// SIMATIC S7-200 project (STEP 7-Micro/WIN), CPU 224XP CN REL 02.01

SYMBOL_TABLE USUARIO1
IN_US            V21.0    // señal de activacion obtenida de la U de transporte
e_k_1            VD132    // error pasado
u_k_1            VD136    // salida pasada
u_k              VD140    // salida U del compensador
V_p              VD124    // Variable de Proceso
e                VD128    // error, diferencia entre REF y V_p
REF              VD104    // nivel de referencia en cm
p_lead           VD116    // polo de adelanto
z_lead           VD112    // zero de adelanto
Kc               VD108    // ganancia compensador
Ts               VD120    // tiempo de muestreo del compensador
SO               I0.3     // Sensor de Objetos (Detecta la pieza para iniciar la seleccion)
S_I              I0.4     // Sensor de fibra Optica (clasificacion de materiales)
SM               I0.5     // Sensor magnetico (clasificacion de materiales)
S1               I0.7     // Sensor de retorno del cilindro 1
S2               I1.0     // Sensor de retorno del cilindro 2
S3               I1.1     // Sensor de retorno del cilindro 3
SBB1             I1.3     // Pulsador de Marcha
SBB2             I1.2     // Pulsador de Paro
QS               I1.4     // Zeta de emergencia
SA               I1.5     // Selector rotatorio
am               Q0.0     // Motor
KV1              Q0.4     // cilindro neumatico 1
KV2              Q0.5     // cilindro neumatico 2
KV3              Q0.6     // cilindro neumatico 3
HL1              Q0.7     // Lampara de señalizacion amarilla
HL2              Q1.0     // Lampara de señalizacion verde
HL3              Q1.1     // Lampara de señalizacion roja
E0               M0.0     // Estado 0
E1               M0.1     // Estado 1
E2               M0.2     // Estado 2
E3               M0.3     // Estado 3
E4               M0.4     // Estado 4
E5               M0.5     // Estado 5
E6               M0.6     // Estado 6
E7               M0.7     // Estado 7
E8               M1.0     // Estado 8
E9               M1.1     // Estado 9
E10              M1.2     // Estado 10
E11              M1.3     // Estado 11
E12              M1.4     // Estado 12
E13              M1.5     // Estado 13
E14              M1.6     // Estado 14
EM               M1.7     // Variable para paro momentaneo
MOTOR            M2.0     // Variable para activacion o desactivacion del motor
E15              M2.1     // Estado 15
E16              M2.2     // Estado 16
SB1_US           V21.1    // Pulsador de marcha
SB2_US           V21.2    // Pulsador de parada
QS_US            V21.3    // Zeta de emergencia
END_SYMBOL_TABLE

ORGANIZATION_BLOCK PRINCIPAL:OB1
TITLE=UNIDAD DE SELECCION
BEGIN
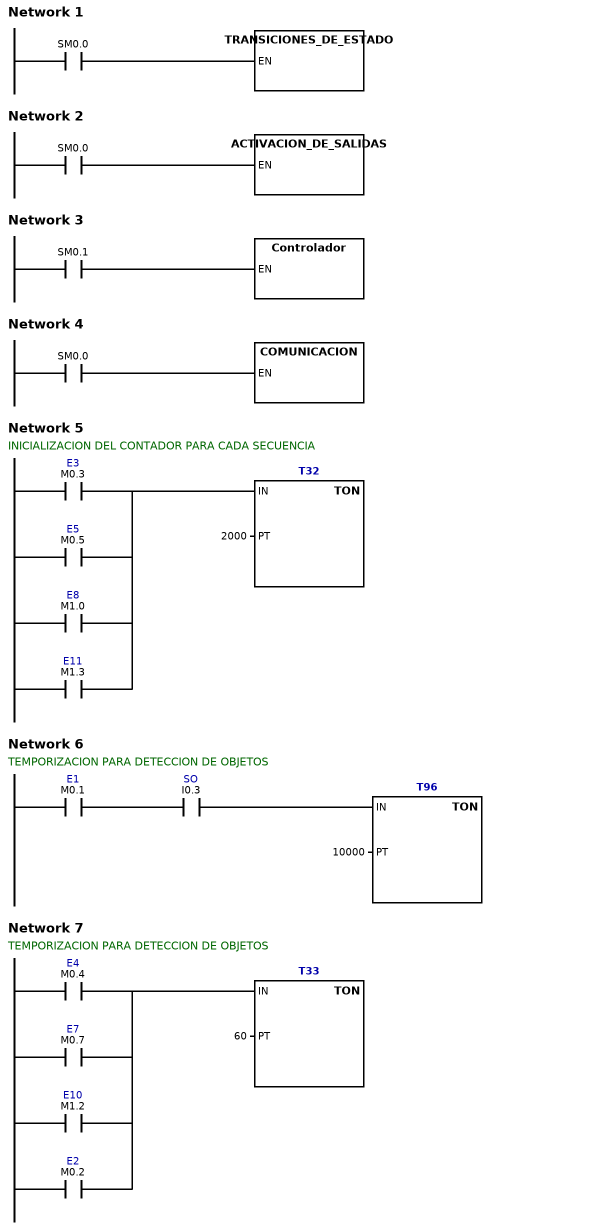
Network 1
LD     SM0.0
CALL   TRANSICIONES_DE_ESTADO:SBR1
Network 2
LD     SM0.0
CALL   ACTIVACION_DE_SALIDAS:SBR2
Network 3
LD     SM0.1
CALL   Controlador:SBR3
Network 4
LD     SM0.0
CALL   COMUNICACION:SBR4
Network 5
// INICIALIZACION DEL CONTADOR PARA CADA SECUENCIA 
LD     E3:M0.3
O      E5:M0.5
O      E8:M1.0
O      E11:M1.3
TON    T32, 2000
Network 6
// TEMPORIZACION PARA DETECCION DE OBJETOS
LD     E1:M0.1
A      SO:I0.3
TON    T96, 10000
Network 7
// TEMPORIZACION PARA DETECCION DE OBJETOS
LD     E4:M0.4
O      E7:M0.7
O      E10:M1.2
O      E2:M0.2
TON    T33, 60
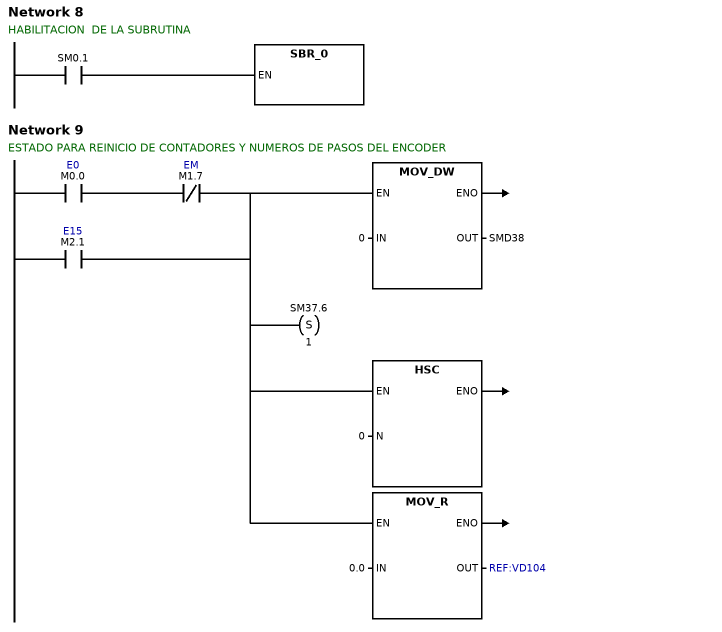
Network 8
// HABILITACION  DE LA SUBRUTINA
LD     SM0.1
CALL   SBR_0:SBR0
Network 9
// ESTADO PARA REINICIO DE CONTADORES Y NUMEROS DE PASOS DEL ENCODER
LD     E0:M0.0
AN     EM:M1.7
O      E15:M2.1
MOVD   0, SMD38
S      SM37.6, 1
HSC    0
MOVR   0.0, REF:VD104
END_ORGANIZATION_BLOCK

SUBROUTINE_BLOCK SBR_0:SBR0
TITLE=COMENTARIOS DE LA SUBRUTINA
BEGIN
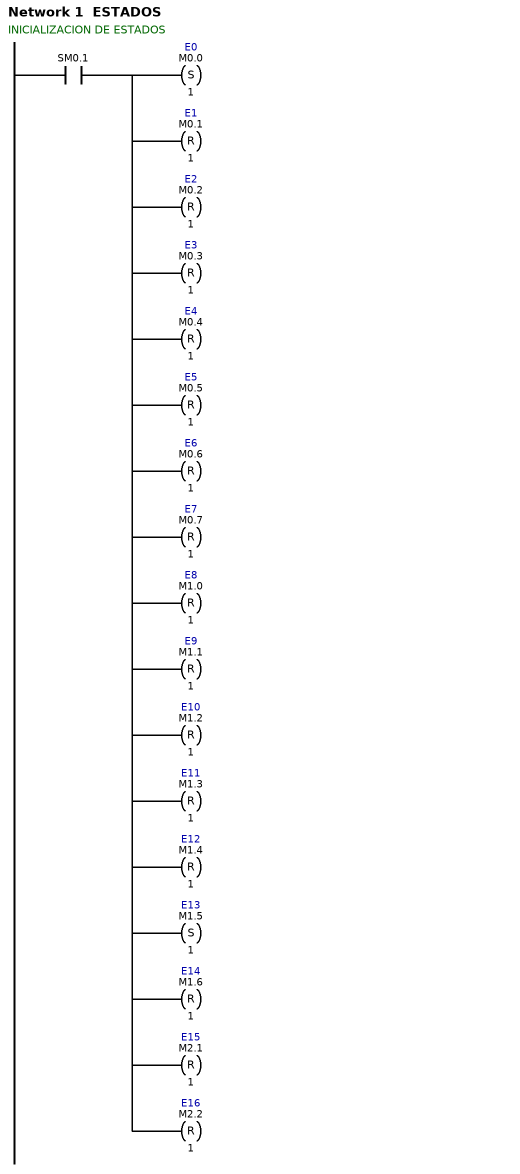
Network 1 // ESTADOS
// INICIALIZACION DE ESTADOS
LD     SM0.1
S      E0:M0.0, 1
R      E1:M0.1, 1
R      E2:M0.2, 1
R      E3:M0.3, 1
R      E4:M0.4, 1
R      E5:M0.5, 1
R      E6:M0.6, 1
R      E7:M0.7, 1
R      E8:M1.0, 1
R      E9:M1.1, 1
R      E10:M1.2, 1
R      E11:M1.3, 1
R      E12:M1.4, 1
S      E13:M1.5, 1
R      E14:M1.6, 1
R      E15:M2.1, 1
R      E16:M2.2, 1
END_SUBROUTINE_BLOCK

SUBROUTINE_BLOCK TRANSICIONES_DE_ESTADO:SBR1
TITLE=TRANSICIONES DE ESTADO
BEGIN
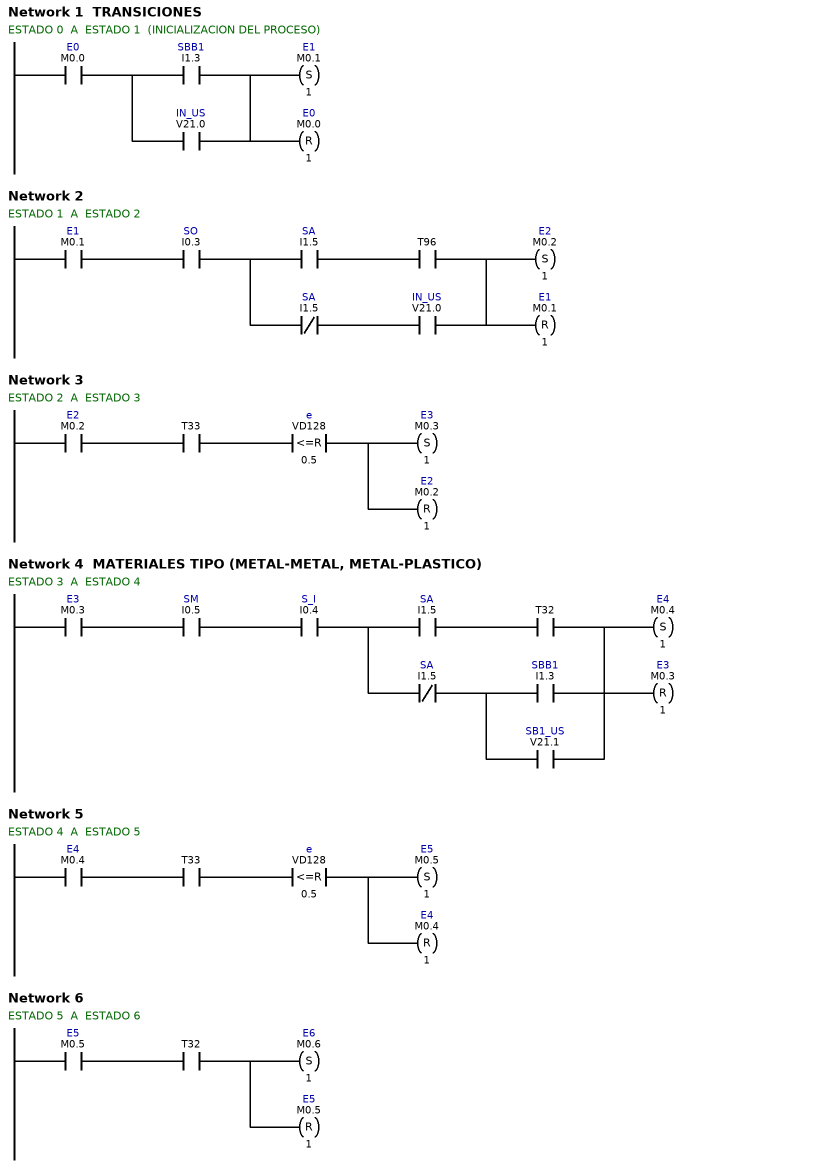
Network 1 // TRANSICIONES
// ESTADO 0  A  ESTADO 1  (INICIALIZACION DEL PROCESO)
LD     E0:M0.0
LD     SBB1:I1.3
O      IN_US:V21.0
ALD
S      E1:M0.1, 1
R      E0:M0.0, 1
Network 2
// ESTADO 1  A  ESTADO 2 
LD     E1:M0.1
A      SO:I0.3
LD     SA:I1.5
A      T96
LDN    SA:I1.5
A      IN_US:V21.0
OLD
ALD
S      E2:M0.2, 1
R      E1:M0.1, 1
Network 3
// ESTADO 2  A  ESTADO 3
LD     E2:M0.2
A      T33
AR<=   e:VD128, 0.5
S      E3:M0.3, 1
R      E2:M0.2, 1
Network 4 // MATERIALES TIPO (METAL-METAL, METAL-PLASTICO)
// ESTADO 3  A  ESTADO 4
LD     E3:M0.3
A      SM:I0.5
A      S_I:I0.4
LD     SA:I1.5
A      T32
LDN    SA:I1.5
LD     SBB1:I1.3
O      SB1_US:V21.1
ALD
OLD
ALD
S      E4:M0.4, 1
R      E3:M0.3, 1
Network 5
// ESTADO 4  A  ESTADO 5
LD     E4:M0.4
A      T33
AR<=   e:VD128, 0.5
S      E5:M0.5, 1
R      E4:M0.4, 1
Network 6
// ESTADO 5  A  ESTADO 6
LD     E5:M0.5
A      T32
S      E6:M0.6, 1
R      E5:M0.5, 1
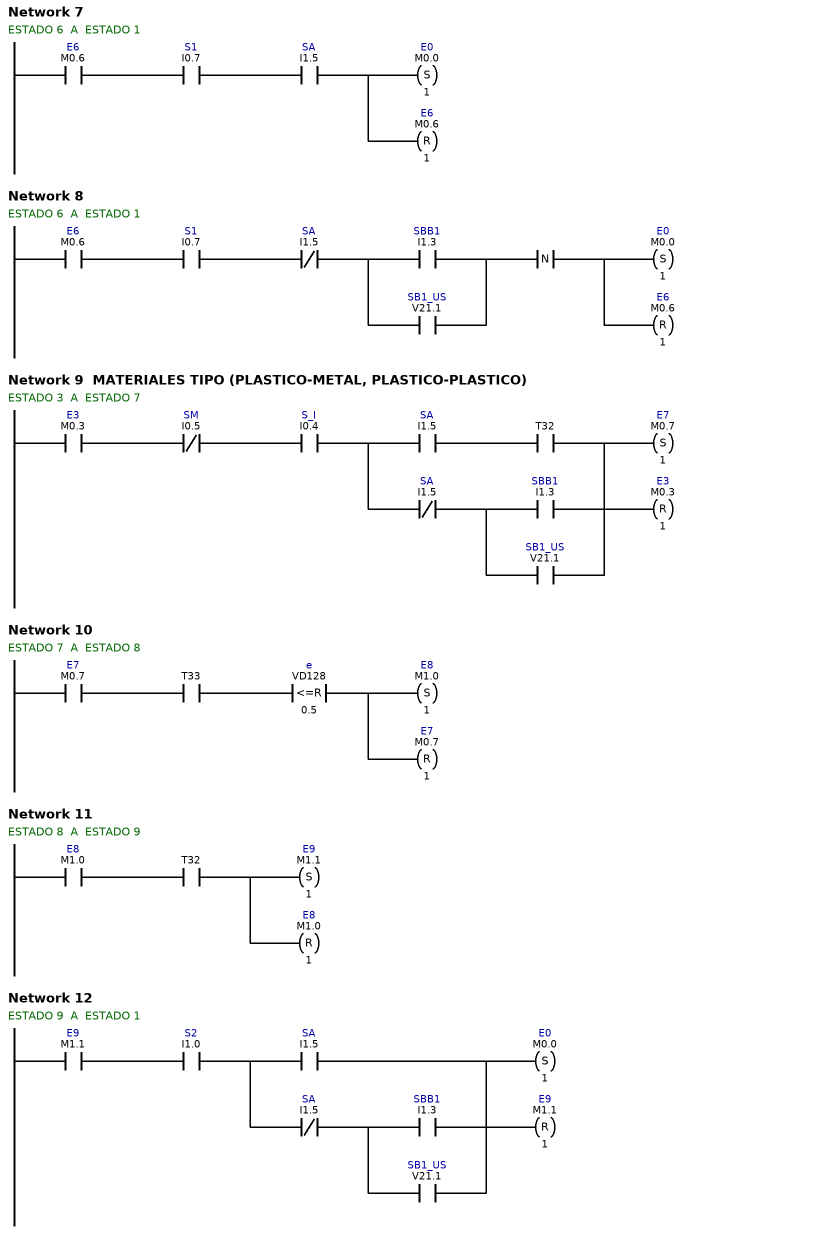
Network 7
// ESTADO 6  A  ESTADO 1
LD     E6:M0.6
A      S1:I0.7
A      SA:I1.5
S      E0:M0.0, 1
R      E6:M0.6, 1
Network 8
// ESTADO 6  A  ESTADO 1
LD     E6:M0.6
A      S1:I0.7
AN     SA:I1.5
LD     SBB1:I1.3
O      SB1_US:V21.1
ALD
ED
S      E0:M0.0, 1
R      E6:M0.6, 1
Network 9 // MATERIALES TIPO (PLASTICO-METAL, PLASTICO-PLASTICO)
// ESTADO 3  A  ESTADO 7
LD     E3:M0.3
AN     SM:I0.5
A      S_I:I0.4
LD     SA:I1.5
A      T32
LDN    SA:I1.5
LD     SBB1:I1.3
O      SB1_US:V21.1
ALD
OLD
ALD
S      E7:M0.7, 1
R      E3:M0.3, 1
Network 10
// ESTADO 7  A  ESTADO 8
LD     E7:M0.7
A      T33
AR<=   e:VD128, 0.5
S      E8:M1.0, 1
R      E7:M0.7, 1
Network 11
// ESTADO 8  A  ESTADO 9
LD     E8:M1.0
A      T32
S      E9:M1.1, 1
R      E8:M1.0, 1
Network 12
// ESTADO 9  A  ESTADO 1
LD     E9:M1.1
A      S2:I1.0
LD     SA:I1.5
LDN    SA:I1.5
LD     SBB1:I1.3
O      SB1_US:V21.1
ALD
OLD
ALD
S      E0:M0.0, 1
R      E9:M1.1, 1
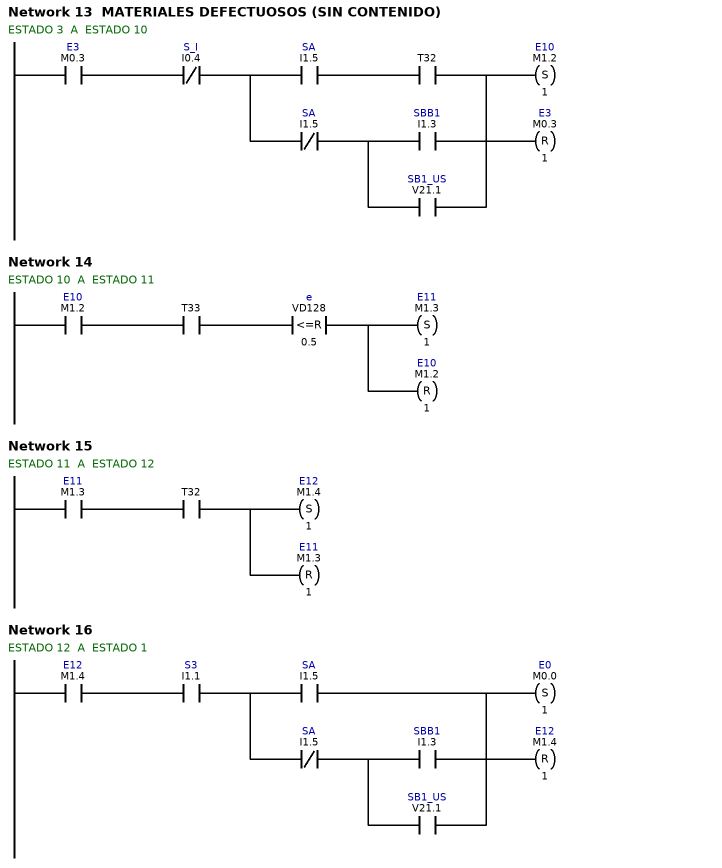
Network 13 // MATERIALES DEFECTUOSOS (SIN CONTENIDO)
// ESTADO 3  A  ESTADO 10 
LD     E3:M0.3
AN     S_I:I0.4
LD     SA:I1.5
A      T32
LDN    SA:I1.5
LD     SBB1:I1.3
O      SB1_US:V21.1
ALD
OLD
ALD
S      E10:M1.2, 1
R      E3:M0.3, 1
Network 14
// ESTADO 10  A  ESTADO 11
LD     E10:M1.2
A      T33
AR<=   e:VD128, 0.5
S      E11:M1.3, 1
R      E10:M1.2, 1
Network 15
// ESTADO 11  A  ESTADO 12
LD     E11:M1.3
A      T32
S      E12:M1.4, 1
R      E11:M1.3, 1
Network 16
// ESTADO 12  A  ESTADO 1
LD     E12:M1.4
A      S3:I1.1
LD     SA:I1.5
LDN    SA:I1.5
LD     SBB1:I1.3
O      SB1_US:V21.1
ALD
OLD
ALD
S      E0:M0.0, 1
R      E12:M1.4, 1
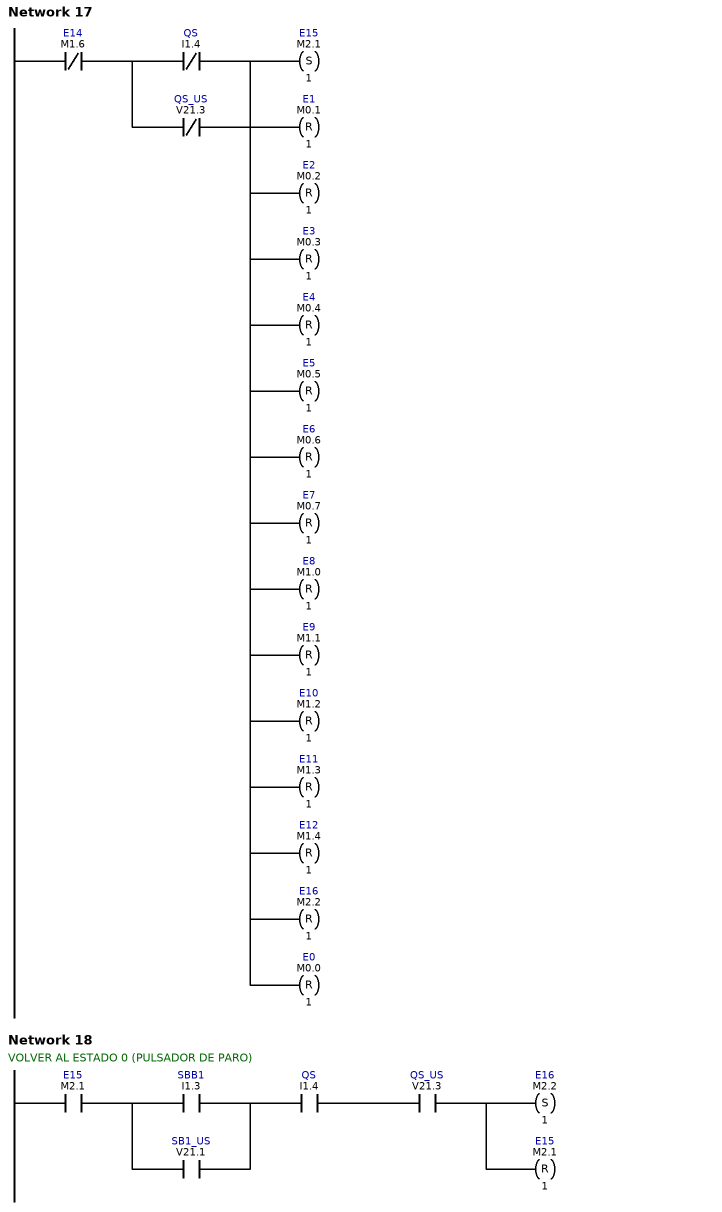
Network 17
LDN    E14:M1.6
LDN    QS:I1.4
ON     QS_US:V21.3
ALD
S      E15:M2.1, 1
R      E1:M0.1, 1
R      E2:M0.2, 1
R      E3:M0.3, 1
R      E4:M0.4, 1
R      E5:M0.5, 1
R      E6:M0.6, 1
R      E7:M0.7, 1
R      E8:M1.0, 1
R      E9:M1.1, 1
R      E10:M1.2, 1
R      E11:M1.3, 1
R      E12:M1.4, 1
R      E16:M2.2, 1
R      E0:M0.0, 1
Network 18
// VOLVER AL ESTADO 0 (PULSADOR DE PARO)
LD     E15:M2.1
LD     SBB1:I1.3
O      SB1_US:V21.1
ALD
A      QS:I1.4
A      QS_US:V21.3
S      E16:M2.2, 1
R      E15:M2.1, 1
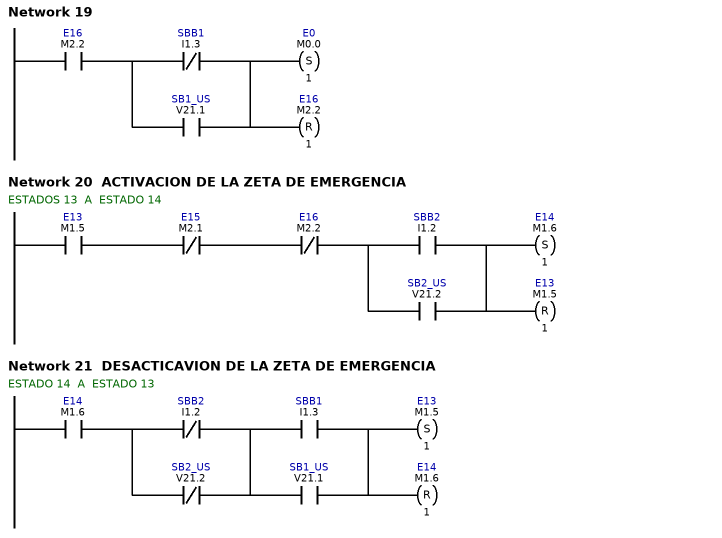
Network 19
LD     E16:M2.2
LDN    SBB1:I1.3
O      SB1_US:V21.1
ALD
S      E0:M0.0, 1
R      E16:M2.2, 1
Network 20 // ACTIVACION DE LA ZETA DE EMERGENCIA
// ESTADOS 13  A  ESTADO 14
LD     E13:M1.5
AN     E15:M2.1
AN     E16:M2.2
LD     SBB2:I1.2
O      SB2_US:V21.2
ALD
S      E14:M1.6, 1
R      E13:M1.5, 1
Network 21 // DESACTICAVION DE LA ZETA DE EMERGENCIA
// ESTADO 14  A  ESTADO 13
LD     E14:M1.6
LDN    SBB2:I1.2
ON     SB2_US:V21.2
ALD
LD     SBB1:I1.3
O      SB1_US:V21.1
ALD
S      E13:M1.5, 1
R      E14:M1.6, 1
Network 22 // Título de segmento
// Comentario de segmento
END_SUBROUTINE_BLOCK

SUBROUTINE_BLOCK ACTIVACION_DE_SALIDAS:SBR2
TITLE=COMENTARIOS DE LA SUBRUTINA
BEGIN
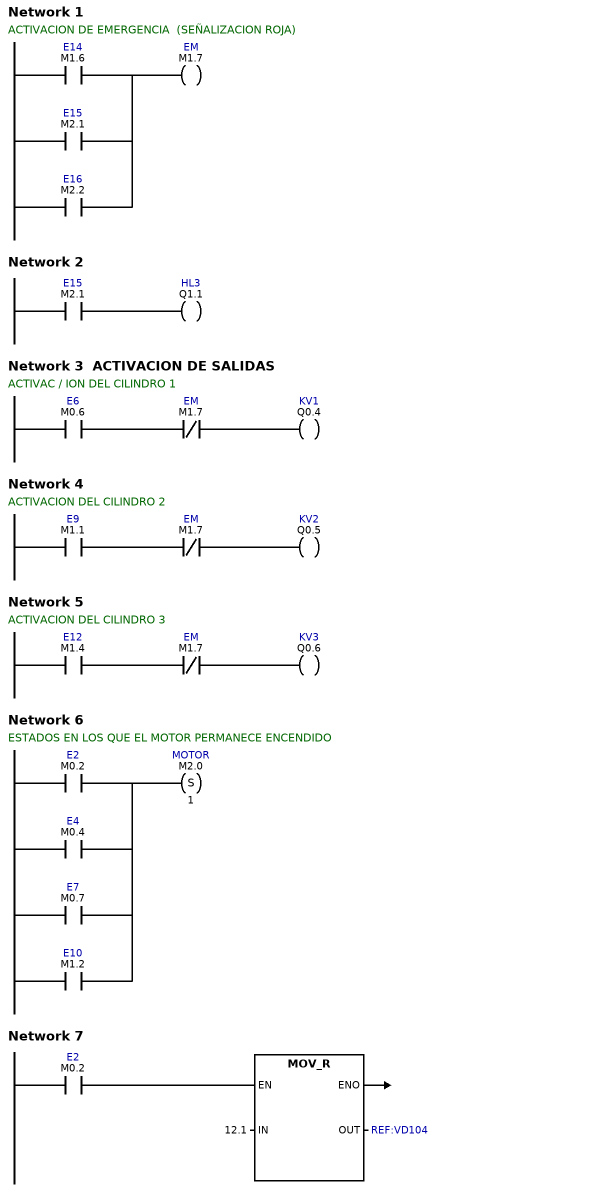
Network 1
// ACTIVACION DE EMERGENCIA  (SEÑALIZACION ROJA)
LD     E14:M1.6
O      E15:M2.1
O      E16:M2.2
=      EM:M1.7
Network 2
LD     E15:M2.1
=      HL3:Q1.1
Network 3 // ACTIVACION DE SALIDAS
// ACTIVAC
// ION DEL CILINDRO 1
LD     E6:M0.6
AN     EM:M1.7
=      KV1:Q0.4
Network 4
// ACTIVACION DEL CILINDRO 2
LD     E9:M1.1
AN     EM:M1.7
=      KV2:Q0.5
Network 5
// ACTIVACION DEL CILINDRO 3
LD     E12:M1.4
AN     EM:M1.7
=      KV3:Q0.6
Network 6
// ESTADOS EN LOS QUE EL MOTOR PERMANECE ENCENDIDO
LD     E2:M0.2
O      E4:M0.4
O      E7:M0.7
O      E10:M1.2
S      MOTOR:M2.0, 1
Network 7
LD     E2:M0.2
MOVR   12.1, REF:VD104
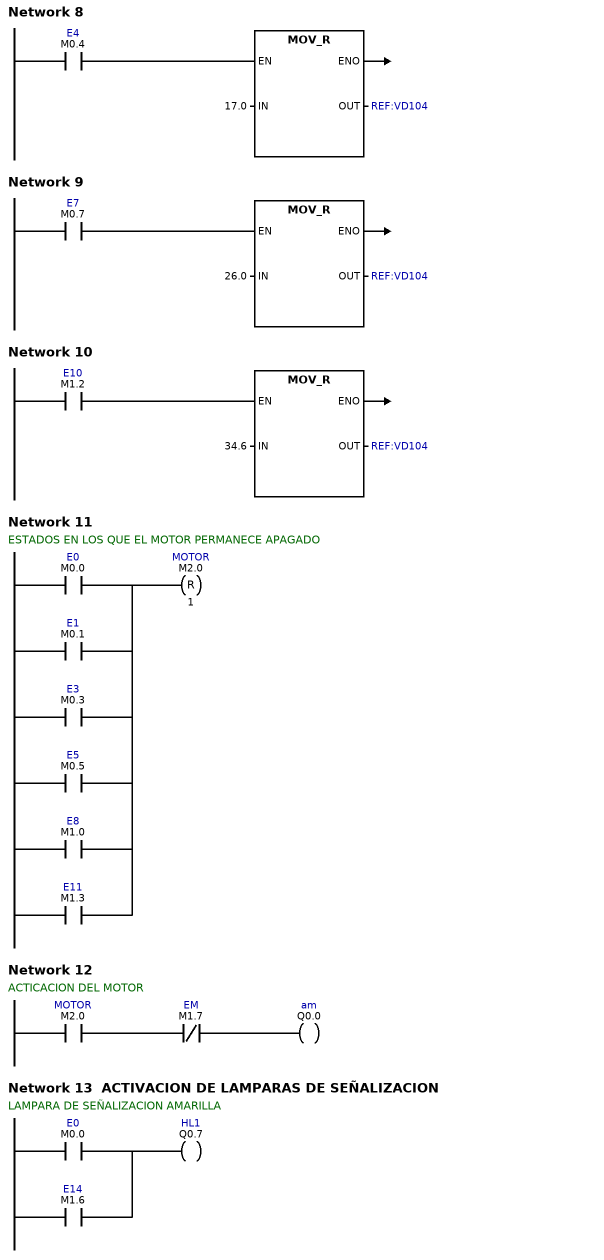
Network 8
LD     E4:M0.4
MOVR   17.0, REF:VD104
Network 9
LD     E7:M0.7
MOVR   26.0, REF:VD104
Network 10
LD     E10:M1.2
MOVR   34.6, REF:VD104
Network 11
// ESTADOS EN LOS QUE EL MOTOR PERMANECE APAGADO
LD     E0:M0.0
O      E1:M0.1
O      E3:M0.3
O      E5:M0.5
O      E8:M1.0
O      E11:M1.3
R      MOTOR:M2.0, 1
Network 12
// ACTICACION DEL MOTOR
LD     MOTOR:M2.0
AN     EM:M1.7
=      am:Q0.0
Network 13 // ACTIVACION DE LAMPARAS DE SEÑALIZACION
// LAMPARA DE SEÑALIZACION AMARILLA
LD     E0:M0.0
O      E14:M1.6
=      HL1:Q0.7
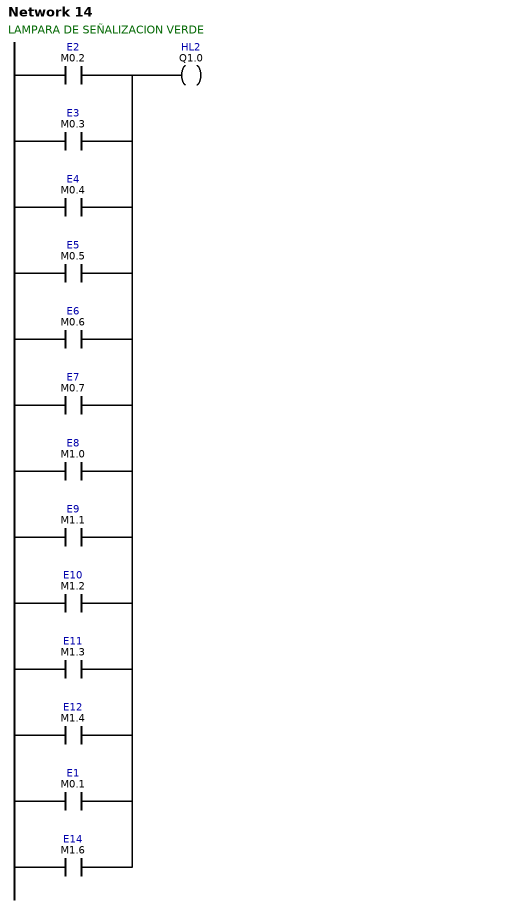
Network 14
// LAMPARA DE SEÑALIZACION VERDE
LD     E2:M0.2
O      E3:M0.3
O      E4:M0.4
O      E5:M0.5
O      E6:M0.6
O      E7:M0.7
O      E8:M1.0
O      E9:M1.1
O      E10:M1.2
O      E11:M1.3
O      E12:M1.4
O      E1:M0.1
O      E14:M1.6
=      HL2:Q1.0
Network 15 // Título de segmento
// Comentario de segmento
END_SUBROUTINE_BLOCK

SUBROUTINE_BLOCK Controlador:SBR3
TITLE=
BEGIN
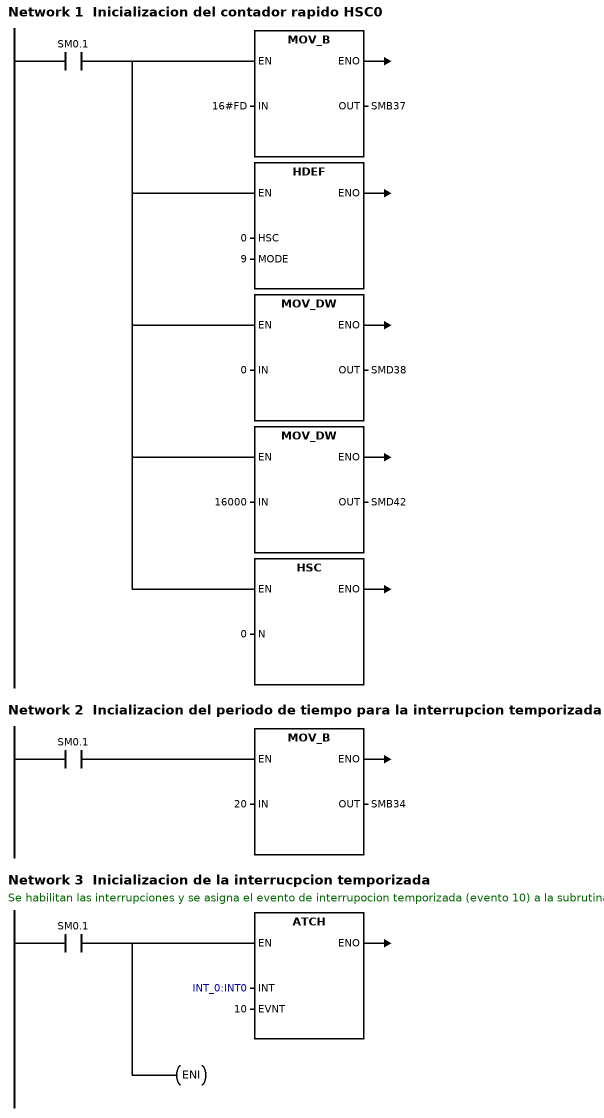
Network 1 // Inicializacion del contador rapido HSC0
LD     SM0.1
MOVB   16#FD, SMB37
HDEF   0, 9
MOVD   0, SMD38
MOVD   16000, SMD42
HSC    0
Network 2 // Incializacion del periodo de tiempo para la interrupcion temporizada
LD     SM0.1
MOVB   20, SMB34
Network 3 // Inicializacion de la interrucpcion temporizada
// Se habilitan las interrupciones y se asigna el evento de interrupocion temporizada (evento 10) a la subrutina de interrupcion INT_0
LD     SM0.1
ATCH   INT_0:INT0, 10
ENI
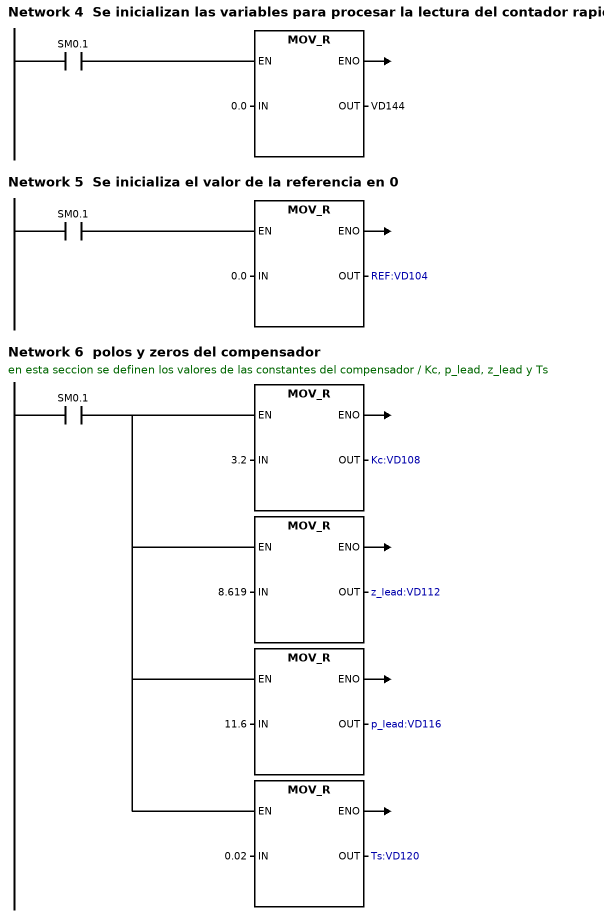
Network 4 // Se inicializan las variables para procesar la lectura del contador rapido HSC0
LD     SM0.1
MOVR   0.0, VD144
Network 5 // Se inicializa el valor de la referencia en 0
LD     SM0.1
MOVR   0.0, REF:VD104
Network 6 // polos y zeros del compensador
// en esta seccion se definen los valores de las constantes del compensador
// Kc, p_lead, z_lead y Ts
LD     SM0.1
MOVR   3.2, Kc:VD108
MOVR   8.619, z_lead:VD112
MOVR   11.6, p_lead:VD116
MOVR   0.02, Ts:VD120
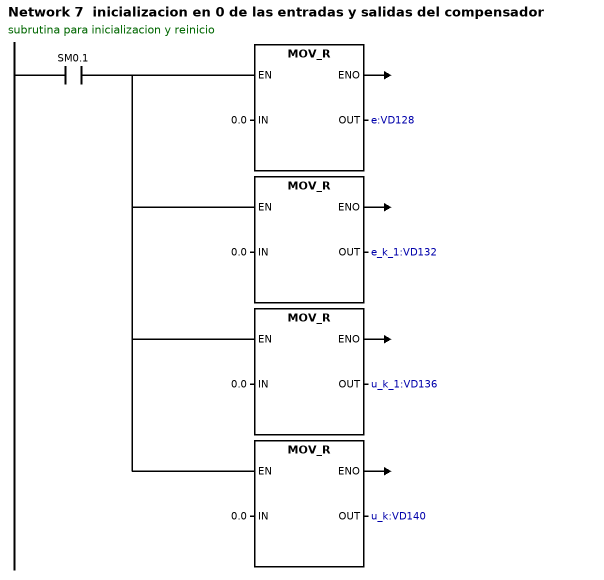
Network 7 // inicializacion en 0 de las entradas y salidas del compensador 
// subrutina para inicializacion y reinicio
LD     SM0.1
MOVR   0.0, e:VD128
MOVR   0.0, e_k_1:VD132
MOVR   0.0, u_k_1:VD136
MOVR   0.0, u_k:VD140
END_SUBROUTINE_BLOCK

SUBROUTINE_BLOCK COMUNICACION:SBR4
TITLE=COMENTARIOS DE LA SUBRUTINA
BEGIN
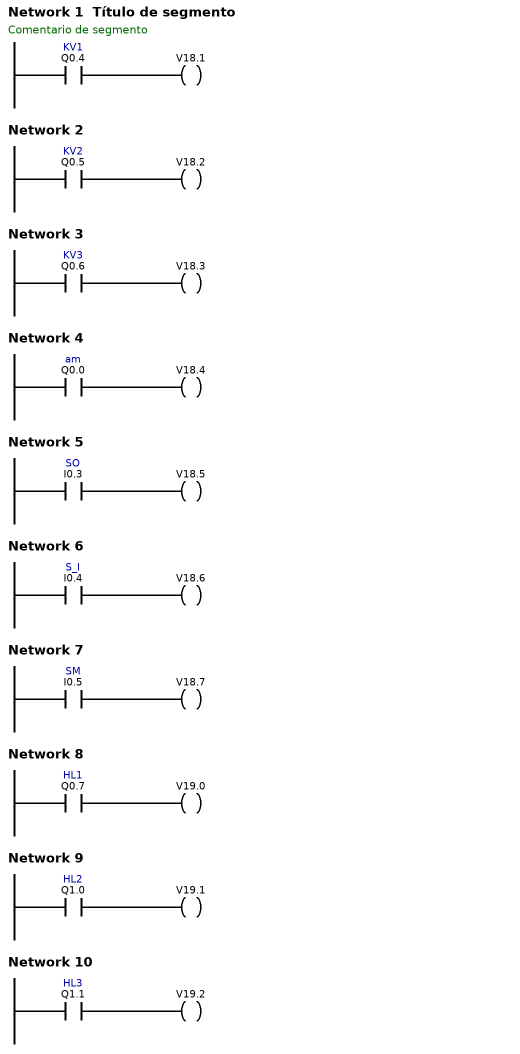
Network 1 // Título de segmento
// Comentario de segmento
LD     KV1:Q0.4
=      V18.1
Network 2
LD     KV2:Q0.5
=      V18.2
Network 3
LD     KV3:Q0.6
=      V18.3
Network 4
LD     am:Q0.0
=      V18.4
Network 5
LD     SO:I0.3
=      V18.5
Network 6
LD     S_I:I0.4
=      V18.6
Network 7
LD     SM:I0.5
=      V18.7
Network 8
LD     HL1:Q0.7
=      V19.0
Network 9
LD     HL2:Q1.0
=      V19.1
Network 10
LD     HL3:Q1.1
=      V19.2
END_SUBROUTINE_BLOCK

INTERRUPT_BLOCK INT_0:INT0
TITLE=
BEGIN
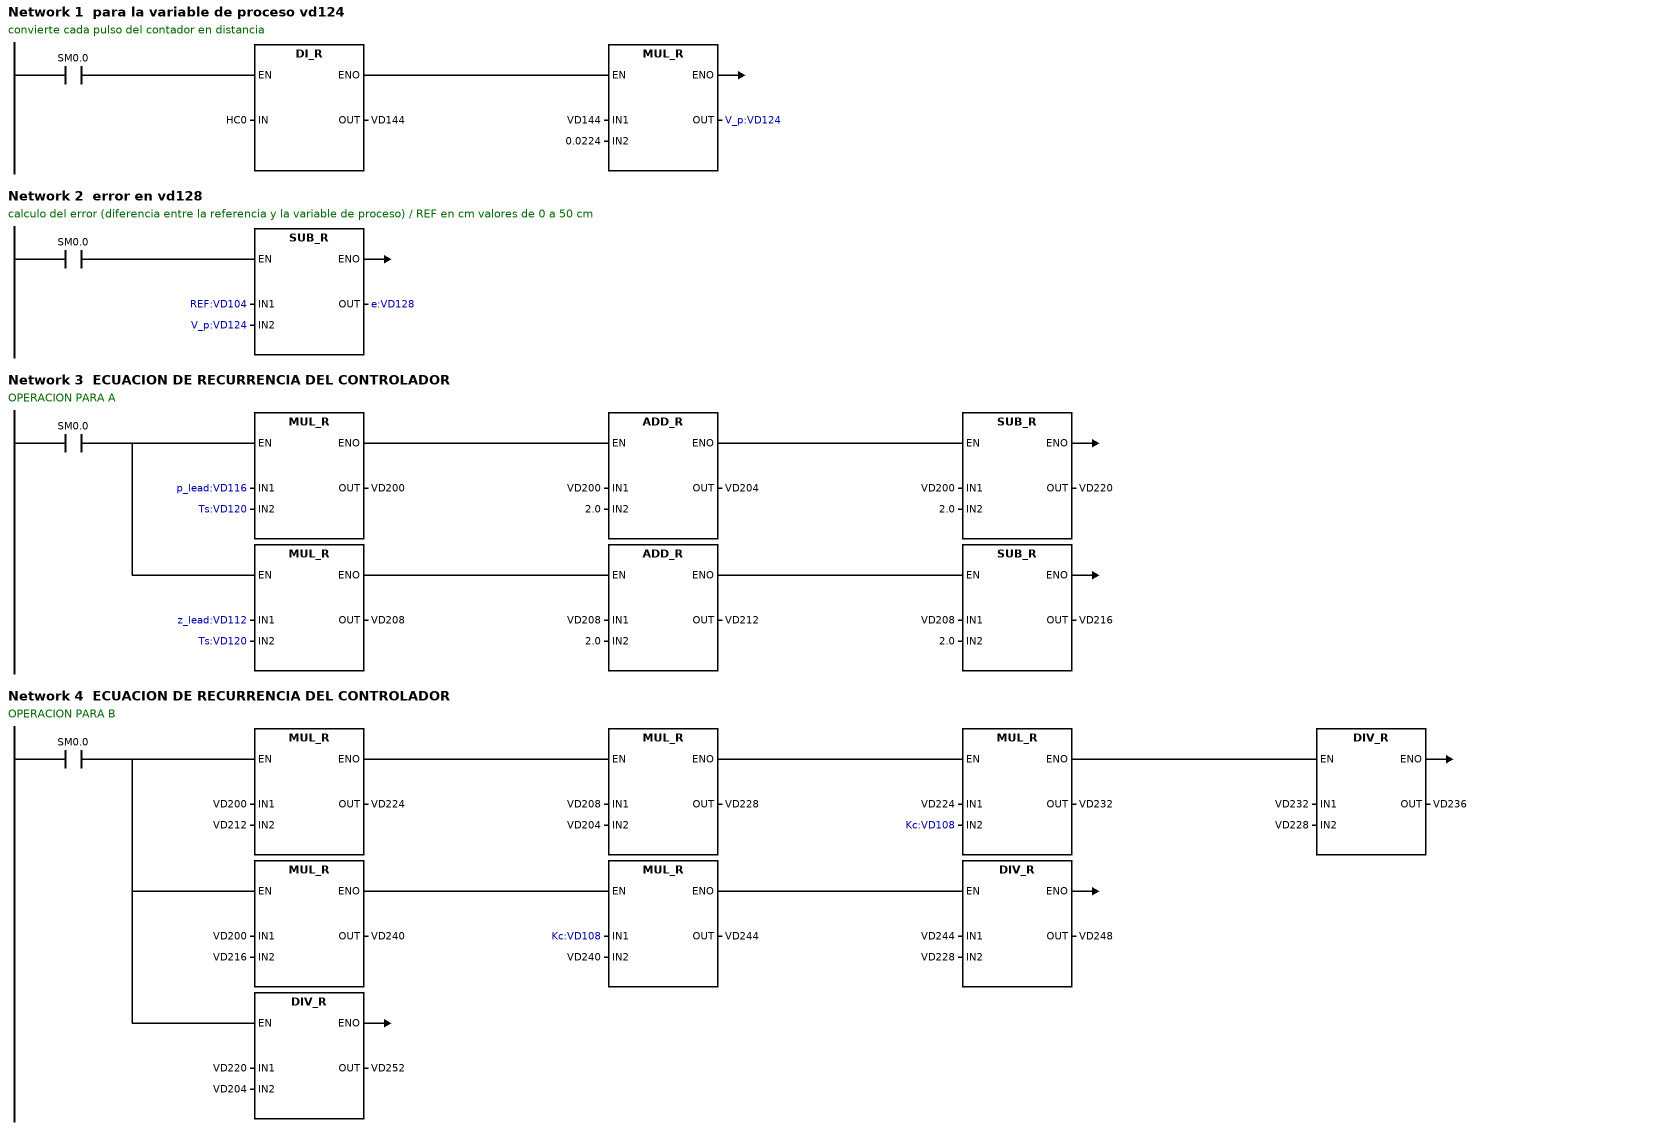
Network 1 // para la variable de proceso vd124
// convierte cada pulso del contador en distancia
LD     SM0.0
DTR    HC0, VD144
AENO
MOVR   VD144, V_p:VD124
*R     0.0224, V_p:VD124
Network 2 // error en vd128
// calculo del error (diferencia entre la referencia y la variable de proceso)
// REF en cm valores de 0 a 50 cm
LD     SM0.0
MOVR   REF:VD104, e:VD128
-R     V_p:VD124, e:VD128
Network 3 // ECUACION DE RECURRENCIA DEL CONTROLADOR
// OPERACION PARA A
LD     SM0.0
LPS
MOVR   p_lead:VD116, VD200
AENO
*R     Ts:VD120, VD200
AENO
MOVR   VD200, VD204
AENO
+R     2.0, VD204
AENO
MOVR   VD200, VD220
-R     2.0, VD220
LPP
MOVR   z_lead:VD112, VD208
AENO
*R     Ts:VD120, VD208
AENO
MOVR   VD208, VD212
AENO
+R     2.0, VD212
AENO
MOVR   VD208, VD216
-R     2.0, VD216
Network 4 // ECUACION DE RECURRENCIA DEL CONTROLADOR
// OPERACION PARA B
LD     SM0.0
LPS
MOVR   VD200, VD224
AENO
*R     VD212, VD224
AENO
MOVR   VD208, VD228
AENO
*R     VD204, VD228
AENO
MOVR   VD224, VD232
AENO
*R     Kc:VD108, VD232
AENO
MOVR   VD232, VD236
/R     VD228, VD236
LRD
MOVR   VD200, VD240
AENO
*R     VD216, VD240
AENO
MOVR   Kc:VD108, VD244
AENO
*R     VD240, VD244
AENO
MOVR   VD244, VD248
/R     VD228, VD248
LPP
MOVR   VD220, VD252
/R     VD204, VD252
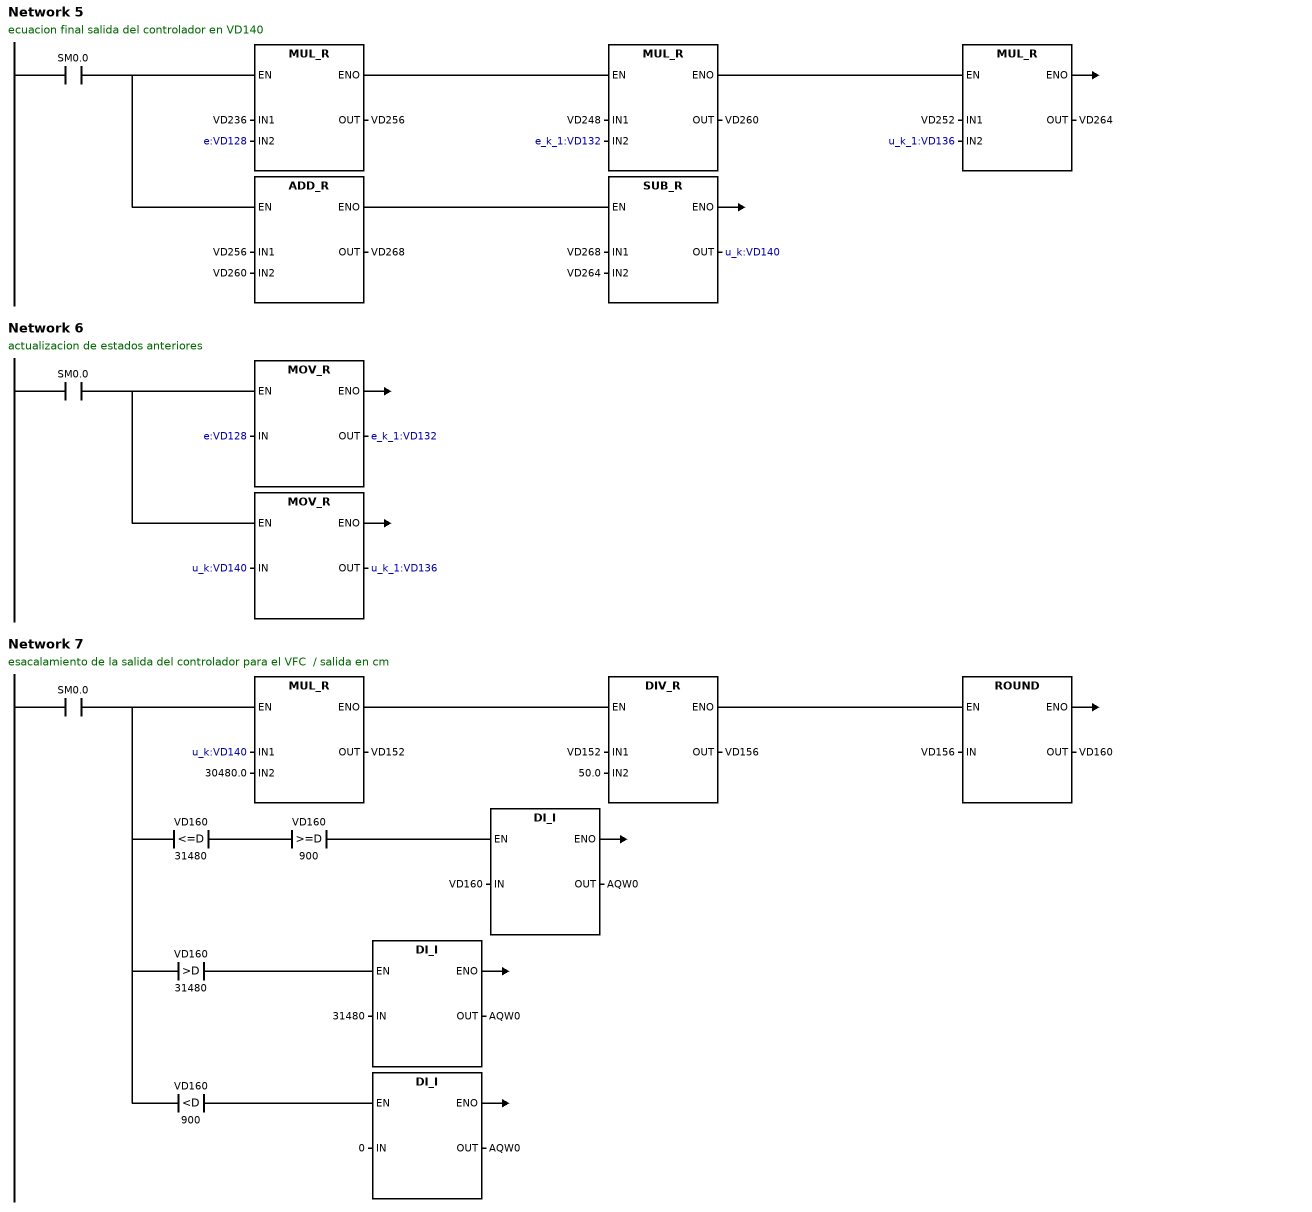
Network 5
// ecuacion final salida del controlador en VD140
LD     SM0.0
LPS
MOVR   VD236, VD256
AENO
*R     e:VD128, VD256
AENO
MOVR   VD248, VD260
AENO
*R     e_k_1:VD132, VD260
AENO
MOVR   VD252, VD264
*R     u_k_1:VD136, VD264
LPP
MOVR   VD256, VD268
AENO
+R     VD260, VD268
AENO
MOVR   VD268, u_k:VD140
-R     VD264, u_k:VD140
Network 6
// actualizacion de estados anteriores
LD     SM0.0
MOVR   e:VD128, e_k_1:VD132
MOVR   u_k:VD140, u_k_1:VD136
Network 7
// esacalamiento de la salida del controlador para el VFC 
// salida en cm
LD     SM0.0
LPS
MOVR   u_k:VD140, VD152
AENO
*R     30480.0, VD152
AENO
MOVR   VD152, VD156
AENO
/R     50.0, VD156
AENO
ROUND  VD156, VD160
LRD
AD<=   VD160, 31480
AD>=   VD160, 900
DTI    VD160, AQW0
LRD
AD>    VD160, 31480
DTI    31480, AQW0
LPP
AD<    VD160, 900
DTI    0, AQW0
END_INTERRUPT_BLOCK
